Fanuc KAREL source: kb00073.KL

-- PROVISIONAL review KL for V1013-1; original PC SHA256 09e2696ce7e7b16143c1edcba9a2097e707ad82cc72942693f6f0620e4ae3fe4
-- Incomplete behavior may be omitted. Consult companion uncertainty JSON. Do not deploy.
PROGRAM KB00073
%NOLOCKGROUP
BEGIN
  -- UNRESOLVED_PC offsets 5-12; opcodes 9D,23
  -- UNRESOLVED_PC offsets 17-26; opcodes 3F,75
  -- UNRESOLVED_PC offsets 31-49; opcodes 27,22,22,2A,31
  -- UNRESOLVED_PC offsets 54-58; opcodes 7F
END KB00073
